// Function block for calculating the substraction of two values
FUNCTION_BLOCK FB_Diff
VAR_INPUT
	var1: UINT;    // variable 1
	var2: UINT;    // variable 2
END_VAR
VAR_OUTPUT
	result : UINT; // result
END_VAR

// Calculation of the substration of two values;
result := var1 - var2;

END_FUNCTION_BLOCK

(* stored: Version 1.1.0.1, ProductVersion 3.1.4026.18
   POU FB_Diff: Id {f3285fee-2279-46b8-82c0-7c9368e56014}, SpecialFunc None *)
